(*
SPDX-FileCopyrightText: c 2026 Oleksandr Tiutyk <trofimich@gmail.com>
SPDX-License-Identifier: MIT
License: https://opensource.org/license/mit
*)

(*!
<summary>Checks exceptions from each hook in both TryCreate paths and writer reset on reuse.</summary>
<description>
Owns persistent native serializer state and any payload buffers used by this case.
Run from one task at a stable address. The caller provides task-boundary exception cleanup.
</description>
*)

{attribute 'no_assign'}
{attribute 'no_explicit_call' := 'do not call this function block directly'}
FUNCTION_BLOCK AutomaticJsonCallbackContainmentAndReuseTest EXTENDS TOF_Testing.SingleCycleTest
VAR_STAT
	{attribute 'hide'}
	_ClassName : STRING := __POUNAME();
END_VAR
VAR
	_Serializer : TOF_JSON.AutomaticJsonSerializer;
	_Extender : JsonExtenderProbe;
	_Source : JSON_TEST_VALUE;
	_Json : TOF_Core.JSON_DOCUMENT;
END_VAR

(*!
<summary>Checks exceptions from each hook in both TryCreate paths and writer reset on reuse.</summary>
*)
METHOD PROTECTED ExecuteTest
VAR
	i : INT;
	sourceInfo : __SYSTEM.VAR_INFO;
	success : BOOL;
	leaked : BOOL;
	jsonSize : UDINT;
	expectedJson : STRING(40) := '[{"Number":42,"Ready":true}]';
END_VAR
_Source.Number := 42;
_Source.Ready := TRUE;

_Json := '';

_Extender.Reset();

sourceInfo := __VARINFO(_Source);

FOR i := 0 TO 3 DO
	_Extender.Reset();
	_Extender.ThrowAtStart := (i MOD 2) = 0;
	_Extender.ThrowAtFinish := NOT _Extender.ThrowAtStart;
	leaked := FALSE;

	__TRY
		IF i < 2 THEN
			success := _Serializer.TrySerialize(
				sourceStructure := _Source,
				extender := _Extender,
				targetJson := _Json,
				jsonSize => jsonSize
			);
		ELSE
			success := _Serializer.TrySerializeByVarInfo(
				sourceStructureVarInfo := sourceInfo,
				sourceStructureAddress := ADR(_Source),
				extender := _Extender,
				targetJson := _Json,
				jsonSize => jsonSize
			);
		END_IF
	__CATCH
		leaked := TRUE;
	__ENDTRY

	Assert.ThatBool(
		actual := leaked,
		message := "Callback exception must not escape Try"
	).IsFalse();
	Assert.ThatBool(
		actual := success,
		message := "Each callback exception must fail Try"
	).IsFalse();
	Assert.ThatUDInt(
		actual := _Extender.StartCount,
		message := "Start must be observed"
	).ToBe(expected := 1);

	IF _Extender.ThrowAtStart THEN
		Assert.ThatUDInt(
			actual := _Extender.FinishCount,
			message := "Failed start must skip finish"
		).ToBe(expected := 0);
	ELSE
		Assert.ThatUDInt(
			actual := _Extender.FinishCount,
			message := "Finish failure must be observed"
		).ToBe(expected := 1);
	END_IF

	_Extender.Reset();
	success := _Serializer.TrySerialize(
		sourceStructure := _Source,
		extender := _Extender,
		targetJson := _Json,
		jsonSize => jsonSize
	);
	Assert.ThatBool(
		actual := success,
		message := "Writer must be reusable after either callback failure"
	).IsTrue();
	Assert.That(
		actual := _Json,
		message := "Reuse must discard the previous partial document"
	).ToBe(expected := expectedJson);
END_FOR
END_METHOD

(*!
<summary>Restores the fixture before the runner publishes the result.</summary>
<description>
Also runs after an unexpected exception interrupts the case.
</description>
*)
METHOD PROTECTED AfterTest
_Extender.Reset();
END_METHOD

//! <summary>Borrows the concrete class name. Callers must not modify it.</summary>
{attribute 'monitoring' := 'call'}
PROPERTY ClassName : REFERENCE TO STRING
GET
ClassName REF= _ClassName;
END_GET
END_PROPERTY

//! <summary>Borrows the compiler-initialized namespace name. Callers must not modify it.</summary>
{attribute 'monitoring' := 'call'}
PROPERTY NamespaceName : REFERENCE TO STRING
GET
NamespaceName REF= CurrentNamespace.Name;
END_GET
END_PROPERTY

//! <summary>Reports the concrete instance size in bytes.</summary>
{attribute 'monitoring' := 'call'}
PROPERTY SelfSize : ULINT
GET
SelfSize := XSIZEOF(THIS^);
END_GET
END_PROPERTY

END_FUNCTION_BLOCK

(* stored: Version 1.1.0.1
   POU AutomaticJsonCallbackContainmentAndReuseTest: Id {2ef77c8e-fc0e-4239-93f0-783a5ba72746}, SpecialFunc None
   Method ExecuteTest: Id {42b1888a-73c7-4b77-9f22-f04861008ccd}
   Method AfterTest: Id {7be871cc-6d90-4466-aac8-99815b41b91d}
   Property ClassName: Id {7dcef803-7878-4b0f-813f-bc54a216edac}
   Get Get: Id {20160fed-aea9-4cc5-abfd-902b93e464f2}
   Property NamespaceName: Id {52966b5c-fef2-4be1-8751-670c78a7937a}
   Get Get: Id {4ced5b63-cac6-4ccf-adf0-82c693b9c2f5}
   Property SelfSize: Id {32318eaf-9849-4022-a24e-0ab9979be9e3}
   Get Get: Id {9916e9bc-83be-46b3-9c12-50cba1840f2e} *)
